Fanuc KAREL source: KX00004.KL

PROGRAM KX00004
%NOLOCKGROUP
VAR
  I: INTEGER
  J: INTEGER
  B: BOOLEAN
  F: FILE
  S: STRING[80]
  P: XYZWPR
BEGIN
  OPEN FILE F ('R', 'MD:KFSAMPLE.DT')
  READ F (I)
  CLOSE FILE F
END KX00004
